(* Logix 5000 project; controller Test vendor 1 type 14 code 167 rev 35.11; software revision 35.00 *)

TASK MainTask (continuous, watchdog 500 ms) : MainProgram

MODULES
   Local : vendor 1 type 14 code 167 (ICP 0, rev 35.11)
END_MODULES

TYPE CMoDateTime :   // Date and Time Structure
STRUCT
   RawDateTime : DINT[7];   // Platform-native wall clock data
   Year : DINT;
   Month : DINT;   // 1-12
   Day : DINT;   // 1-31
   Hour : DINT;   // 0-23
   Minute : DINT;   // 0-59
   Second : DINT;   // 0-59
   MicroSecond : DINT;   // 0-999999
   IsLocal : BOOL;   // TRUE = local time, FALSE = UTC
END_STRUCT
END_TYPE

TYPE CMoDateTimeString :   // HMI-Readable Date/Time Strings
STRUCT
   TimeString : CMoString28;   // HH:MM:SS
   DateString : CMoString28;   // YYYY-MM-DD
   HMIString : CMoString28;   // YYYY-MM-DD HH:MM:SS
END_STRUCT
END_TYPE

TYPE CMoFramework :   // Shared System Context - one per PLC
STRUCT
   AnyAudibleOn : BOOL;   // Audible alarm active
   AnyAudibleOnLastScan : BOOL;   // Scratch
   AnyAlarmActive : BOOL;   // Alarm active
   AnyAlarmActiveLastScan : BOOL;   // Scratch
   AnyWarningActive : BOOL;   // Warning active
   AnyWarningActiveLastScan : BOOL;   // Scratch
   AnyFaultActive : BOOL;   // Fault active
   AnyFaultActiveLastScan : BOOL;   // Scratch
   AnyCriticalActive : BOOL;   // Critical active
   AnyCriticalActiveLastScan : BOOL;   // Scratch
   AnySimulationOn : BOOL;   // Sim active
   AnySimulationOnLastScan : BOOL;   // Scratch
   AnyHandOn : BOOL;   // Hand active
   AnyHandOnLastScan : BOOL;   // Scratch
   SilenceCmd : BOOL;   // HMI silence (momentary)
   GlobalAlmRstCmd : BOOL;   // HMI global reset (momentary)
   GlobalAlmRstEn : BOOL;   // Enable global reset
   SimulationEnabled : BOOL;   // Master sim enable
   EmulationEnabled : BOOL;   // Emulated controller
   MaintenanceEnabled : BOOL;   // Enables Hand mode
   Tick100ms : BOOL;   // 100ms tick
   Tick1s : BOOL;   // 1s tick
   Tick10s : BOOL;   // 10s tick
   Blink100ms : BOOL;   // 100ms blinker
   Blink250ms : BOOL;   // 250ms blinker
   Blink500ms : BOOL;   // 500ms blinker
   Blink1s : BOOL;   // 1s blinker
   Blink2s : BOOL;   // 2s blinker
   InhibitAlarms : BOOL;   // Corporate alarm inhibit
   AlwaysTrue : BOOL;   // Constant TRUE
   AlwaysFalse : BOOL;   // Constant FALSE
   ApplicationCount : DINT;   // AOI instance count
   AlarmCount : INT;   // Active alarm count
   TempAlarmCount : INT;   // Scratch
   FreeRunningTimer : DINT;   // Free-running ms counter
   LastRandomSeed : DINT;   // Random seed
   Random : REAL;   // Random 0.0-1.0
   CycleTime : REAL;   // Scan time (ms)
   InhibitAlarmGroups : DINT[16];   // Per-group inhibit (512 groups)
   CurrentUTCDateTime : CMoDateTime;   // UTC time
   CurrentLocalDateTime : CMoDateTime;   // Local time
   CurrentUTCString : CMoDateTimeString;   // UTC strings
   CurrentLocalString : CMoDateTimeString;   // Local strings
   NotUsedDI : CMoHALDigitalInput;   // Spare DI
   NotUsedDO : CMoHALDigitalOutput;   // Spare DO
   ModuleStatusMinInterval : DINT;   // ms between module checks
   ModuleStatusRandomDistribution : DINT;   // ms random spread
   ModuleStatusGraceTime : DINT;   // ms before module lost
END_STRUCT
END_TYPE

TYPE CMoHALDigitalInput :   // Digital Input HAL - Business logic reads .Value only
STRUCT
   Input : BOOL;   // Raw hardware input
   QualityInput : BOOL;   // Hardware health (TRUE = good)
   SimInput : BOOL;   // Simulation input (twin/test)
   EnableSimulation : BOOL;   // Enable simulation for this point
   SimulationIsActive : BOOL;   // Computed: EnableSimulation AND Framework.SimulationEnabled
   HandValue : BOOL;   // Manual override value (HMI)
   EnableHand : BOOL;   // Enable hand mode
   HandIsActive : BOOL;   // Computed: EnableHand AND Framework.MaintenanceEnabled
   Value : BOOL;   // THE OUTPUT: conditioned, filtered, mode-selected
   Inverted : BOOL;   // Invert input polarity
   BadQualityValue : BOOL;   // Value when quality is bad
   EnableDelay : BOOL;   // Enable debounce filtering
   IsSpare : BOOL;   // Mark as spare
   InFilterOnTimeMsec : DINT;   // On-delay debounce (ms)
   InFilterOffTimeMsec : DINT;   // Off-delay debounce (ms)
   PointQuality : BOOL;   // Computed quality
   RisingEdge : BOOL;   // One-shot on Value 0->1
   FallingEdge : BOOL;   // One-shot on Value 1->0
   Name : CMoString28;   // Human-readable tag name
END_STRUCT
END_TYPE

TYPE CMoHALDigitalOutput :   // Digital Output HAL - Business logic writes .Value
STRUCT
   Output : BOOL;   // Physical output
   QualityInput : BOOL;   // Hardware health (TRUE = good)
   SimOutput : BOOL;   // Shadow output for twin
   EnableSimulation : BOOL;   // Enable simulation
   SimulationIsActive : BOOL;   // Computed
   HandValue : BOOL;   // Manual override value
   EnableHand : BOOL;   // Enable hand mode
   HandIsActive : BOOL;   // Computed
   Value : BOOL;   // Business logic command
   Inverted : BOOL;   // Invert output polarity
   BadQualityValue : BOOL;   // Value when quality is bad
   IsSpare : BOOL;   // Mark as spare
   PointQuality : BOOL;   // Computed quality
   Name : CMoString28;   // Human-readable tag name
END_STRUCT
END_TYPE

TYPE CMoInterlock :   // Interlock: 16 AND conditions, first-out, per-condition bypass
STRUCT
   PointCount : INT;   // Number of active conditions (1-16)
   Condition : BOOL[32];   // Condition inputs
   Bypass : BOOL[32];   // Per-condition bypass (HMI)
   OK : BOOL;   // All conditions met or bypassed
   InBypass : BOOL;   // At least one bypassed
   BypassAlarm : BOOL;   // Operating with bypass
   FirstOut : INT;   // First faulted condition index (-1=none)
   ConditionMet : BOOL[32];   // Condition OR bypass
   ConditionFaulted : BOOL[32];   // Failed AND not bypassed
   Name : CMoString28;   // Interlock name
   ConditionName : CMoString28[16];   // Per-condition labels
END_STRUCT
END_TYPE

TYPE CMoString28 :
STRUCT
   LEN : DINT;
   DATA : SINT[28];
END_STRUCT
END_TYPE

ADD_ON_INSTRUCTION CMoAlarm   (* revision 1.0 *)
// Alarm Monitor
// Help:
// Trigger, delay, reset, severity, group inhibit, silencing, occurrence counting.
VAR_IN_OUT
   Framework : CMoFramework; {required}   // System context
END_VAR
VAR_INPUT
   Trigger : BOOL;   // Condition to monitor
   EnableAlarm : BOOL := 1;   // Enable this alarm
   AlarmOnTrue : BOOL := 1;   // Trigger=1 alarms
   AutoReset : BOOL;   // Auto-clear
   Delay : DINT;   // ms before activating
   GroupNo : DINT;   // Alarm group 0-511
   ID : INT;   // Alarm ID 1-9023
   IsWarning : BOOL;   // Warning severity
   IsFault : BOOL;   // Fault severity
   IsCritical : BOOL;   // Critical severity
   EnableAudio : BOOL;   // Enable audible
   SystemResetEnable : BOOL := 1;   // Allow global reset
   Reset : BOOL;   // Manual reset
   Inhibit : BOOL;   // Per-alarm inhibit
   CountPreset : DINT;   // Count threshold
   CountReset : BOOL;   // Reset counter
END_VAR
VAR_OUTPUT
   AlarmActive : BOOL; {access Read Only}   // Alarm is active
   InhibitActive : BOOL; {access Read Only}   // Currently inhibited
   AlarmCount : DINT; {access Read Only}   // Activation count
   CountExceeded : BOOL; {access Read Only}   // Count >= preset
   AlarmSilenced : BOOL; {access Read Only}   // Active but silenced
END_VAR
VAR
   AlarmTimer : FBD_TIMER; {access None}
   IntGroupNo : DINT; {access None}
   IntID : DINT; {access None}
   IntReset : BOOL; {access None}
   TriggerCondition : BOOL; {access None}
   PrevAlarmActive : BOOL; {access None}
END_VAR

ROUTINE Logic   (* structured text *)
   // =============================================================================
   // CMoAlarm — Alarm Monitor
   // CMo Library v1.0
   // =============================================================================
   // Monitors a trigger condition and manages alarm lifecycle.
   // Supports configurable trigger polarity, delay before activation,
   // auto/manual reset, occurrence counting with threshold,
   // severity classification (Warning/Fault/Critical), group-based
   // inhibit, and HMI silencing.
   // =============================================================================
   
   IF GroupNo >= 0 AND GroupNo <= 511 THEN IntGroupNo := GroupNo; ELSE IntGroupNo := 0; END_IF;
   IF ID >= 1 AND ID <= 9023 THEN IntID := ID; ELSE IntID := 0; END_IF;
   IF CountReset THEN AlarmCount := 0; CountReset := 0; END_IF;
   InhibitActive := NOT EnableAlarm OR Inhibit OR Framework.InhibitAlarms;
   IntReset := AutoReset OR Reset OR (SystemResetEnable AND Framework.GlobalAlmRstEn AND Framework.GlobalAlmRstCmd);
   IF AlarmOnTrue THEN TriggerCondition := Trigger; ELSE TriggerCondition := NOT Trigger; END_IF;
   
   IF IntID <> 0 THEN
       AlarmTimer.PRE := Delay;
       AlarmTimer.TimerEnable := (NOT InhibitActive AND TriggerCondition) OR (AlarmActive AND NOT IntReset);
       TONR(AlarmTimer);
       AlarmActive := AlarmTimer.DN;
       IF NOT AlarmTimer.TimerEnable THEN
           AlarmTimer.Reset := 1; TONR(AlarmTimer); AlarmTimer.Reset := 0;
       END_IF;
   ELSE
       AlarmActive := 0;
   END_IF;
   
   IF AlarmActive AND NOT PrevAlarmActive THEN AlarmCount := AlarmCount + 1; END_IF;
   IF AlarmActive THEN
       IF Framework.SilenceCmd OR AlarmSilenced THEN AlarmSilenced := 1; END_IF;
   ELSE AlarmSilenced := 0;
   END_IF;
   
   IF AlarmActive THEN
       Framework.TempAlarmCount := Framework.TempAlarmCount + 1;
       Framework.AnyAlarmActiveLastScan := 1;
       IF NOT AlarmSilenced THEN
           IF EnableAudio THEN Framework.AnyAudibleOnLastScan := 1; END_IF;
           IF IsWarning THEN Framework.AnyWarningActiveLastScan := 1; END_IF;
           IF IsFault THEN Framework.AnyFaultActiveLastScan := 1; END_IF;
           IF IsCritical THEN Framework.AnyCriticalActiveLastScan := 1; END_IF;
       END_IF;
   END_IF;
   
   IF CountPreset > 0 AND AlarmCount >= CountPreset THEN CountExceeded := 1; ELSE CountExceeded := 0; END_IF;
   Reset := 0;
   PrevAlarmActive := AlarmActive;
END_ROUTINE
END_ADD_ON_INSTRUCTION

ADD_ON_INSTRUCTION CMoDateTimeToString   (* revision 1.0 *)
// Format DateTime for HMI Display
// Help:
// Converts CMoDateTime into zero-padded strings.
VAR_IN_OUT
   DateTime : CMoDateTime; {required}   // Input DateTime
   DateTimeString : CMoDateTimeString; {required}   // Output formatted strings
END_VAR
VAR
   sYear : CMoString28; {access None}
   sMonth : CMoString28; {access None}
   sDay : CMoString28; {access None}
   sHour : CMoString28; {access None}
   sMinute : CMoString28; {access None}
   sSecond : CMoString28; {access None}
   sTemp : CMoString28; {access None}
   sZero : CMoString28; {access None}
   sColon : CMoString28; {access None}
   sDash : CMoString28; {access None}
   sBlank : CMoString28; {access None}
END_VAR

ROUTINE Logic   (* structured text *)
   // =============================================================================
   // CMoDateTimeToString — Format DateTime for HMI Display
   // CMo Library v1.0
   // =============================================================================
   // Converts CMoDateTime fields into zero-padded human-readable strings:
   //   TimeString: "HH:MM:SS"
   //   DateString: "YYYY-MM-DD"
   //   HMIString:  "YYYY-MM-DD HH:MM:SS"
   //
   // Uses DTOS for DINT-to-string conversion.
   // =============================================================================
   
   DTOS(DateTime.Year, sYear);
   sZero := '0';
   sColon := ':';
   sDash := '-';
   sBlank := ' ';
   IF DateTime.Month < 10 THEN
       DTOS(DateTime.Month, sTemp);
       CONCAT(sZero, sTemp, sMonth);
   ELSE
       DTOS(DateTime.Month, sMonth);
   END_IF;
   
   IF DateTime.Day < 10 THEN
       DTOS(DateTime.Day, sTemp);
       CONCAT(sZero, sTemp, sDay);
   ELSE
       DTOS(DateTime.Day, sDay);
   END_IF;
   
   IF DateTime.Hour < 10 THEN
       DTOS(DateTime.Hour, sTemp);
       CONCAT(sZero, sTemp, sHour);
   ELSE
       DTOS(DateTime.Hour, sHour);
   END_IF;
   
   IF DateTime.Minute < 10 THEN
       DTOS(DateTime.Minute, sTemp);
       CONCAT(sZero, sTemp, sMinute);
   ELSE
       DTOS(DateTime.Minute, sMinute);
   END_IF;
   
   IF DateTime.Second < 10 THEN
       DTOS(DateTime.Second, sTemp);
       CONCAT(sZero, sTemp, sSecond);
   ELSE
       DTOS(DateTime.Second, sSecond);
   END_IF;
   
   // Build TimeString: "HH:MM:SS"
   
   CONCAT(sHour, sColon, sTemp);
   CONCAT(sTemp, sMinute, sTemp);
   CONCAT(sTemp, sColon, sTemp);
   CONCAT(sTemp, sSecond, DateTimeString.TimeString);
   
   // Build DateString: "YYYY-MM-DD"
   CONCAT(sYear, sDash, sTemp);
   CONCAT(sTemp, sMonth, sTemp);
   CONCAT(sTemp, sDash, sTemp);
   CONCAT(sTemp, sDay, DateTimeString.DateString);
   
   // Build HMIString: "YYYY-MM-DD HH:MM:SS"
   CONCAT(DateTimeString.DateString, sBlank, sTemp);
   CONCAT(sTemp, DateTimeString.TimeString, DateTimeString.HMIString);
END_ROUTINE
END_ADD_ON_INSTRUCTION

ADD_ON_INSTRUCTION CMoDiffTime   (* revision 1.0 *)
// DateTime Subtraction with Carry Propagation
// Help:
// Computes EndTime - StartTime with carry propagation.
VAR_IN_OUT
   StartTime : CMoDateTime; {required}   // Start time
   EndTime : CMoDateTime; {required}   // End time
   Result : CMoDateTime; {required}   // Difference result
END_VAR
VAR_OUTPUT
   TotalSeconds : DINT; {access Read Only}   // Approximate total seconds
   TotalMicroseconds : DINT; {access Read Only}   // Remainder microseconds
END_VAR
VAR
   a : DINT; {access None}
   y : DINT; {access None}
   m : DINT; {access None}
   jdnStart : DINT; {access None}
   jdnEnd : DINT; {access None}
   diffDays : DINT; {access None}
   diffUs : DINT; {access None}
   diffSec : DINT; {access None}
   diffMin : DINT; {access None}
   diffHr : DINT; {access None}
END_VAR

ROUTINE Logic   (* structured text *)
   // =============================================================================
   // CMoDiffTime — DateTime Subtraction via Julian Day Number
   // CMo Library v1.0 — Rockwell
   // =============================================================================
   // Computes (EndTime - StartTime) using Julian Day Number conversion.
   // Converts both dates to JDN (integer day count), subtracts, then
   // handles sub-day time remainder with borrow propagation.
   //
   // This is mathematically correct for all valid dates regardless of
   // month lengths, leap years, or century boundaries.
   //
   // Usage:
   //   CMoDiffTime(fbDiff, tStart, tEnd, tResult);
   //   elapsed := fbDiff.TotalSeconds;
   // =============================================================================
   
   // JDN for StartTime
   a := (14 - StartTime.Month) / 12;
   y := StartTime.Year + 4800 - a;
   m := StartTime.Month + 12 * a - 3;
   jdnStart := StartTime.Day + (153 * m + 2) / 5 + 365 * y + y / 4 - y / 100 + y / 400 - 32045;
   
   // JDN for EndTime
   a := (14 - EndTime.Month) / 12;
   y := EndTime.Year + 4800 - a;
   m := EndTime.Month + 12 * a - 3;
   jdnEnd := EndTime.Day + (153 * m + 2) / 5 + 365 * y + y / 4 - y / 100 + y / 400 - 32045;
   
   // Day difference
   diffDays := jdnEnd - jdnStart;
   
   // Sub-day difference with borrow propagation
   diffUs := EndTime.MicroSecond - StartTime.MicroSecond;
   IF diffUs < 0 THEN
       diffUs := diffUs + 1000000;
       diffSec := -1;
   ELSE
       diffSec := 0;
   END_IF;
   
   diffSec := diffSec + EndTime.Second - StartTime.Second;
   IF diffSec < 0 THEN
       diffSec := diffSec + 60;
       diffMin := -1;
   ELSE
       diffMin := 0;
   END_IF;
   
   diffMin := diffMin + EndTime.Minute - StartTime.Minute;
   IF diffMin < 0 THEN
       diffMin := diffMin + 60;
       diffHr := -1;
   ELSE
       diffHr := 0;
   END_IF;
   
   diffHr := diffHr + EndTime.Hour - StartTime.Hour;
   IF diffHr < 0 THEN
       diffHr := diffHr + 24;
       diffDays := diffDays - 1;
   END_IF;
   
   // Populate result
   Result.Year := 0;
   Result.Month := 0;
   Result.Day := diffDays;
   Result.Hour := diffHr;
   Result.Minute := diffMin;
   Result.Second := diffSec;
   Result.MicroSecond := diffUs;
   Result.IsLocal := 0;
   
   // Convenience totals
   TotalSeconds := diffSec + (diffMin * 60) + (diffHr * 3600) + (diffDays * 86400);
   TotalMicroseconds := diffUs;
END_ROUTINE
END_ADD_ON_INSTRUCTION

ADD_ON_INSTRUCTION CMoDigitalInput   (* revision 1.0 *)
// Digital Input Signal Conditioning
// Help:
// Mode select, inversion, debounce, quality gating, edge detection. Reads .Value only.
VAR_IN_OUT
   HAL : CMoHALDigitalInput; {required}   // HAL Interface
END_VAR
VAR_INPUT
   DeviceInput : BOOL; {required}   // Raw hardware input
   QualityInput : BOOL; {required}   // Module health
END_VAR
VAR_IN_OUT
   Framework : CMoFramework; {required}   // System context
END_VAR
VAR
   ConditionedInput : BOOL; {access None}
   DebouncedValue : BOOL; {access None}
   OnDelayTimer : FBD_TIMER; {access None}
   OffDelayTimer : FBD_TIMER; {access None}
   PrevValue : BOOL; {access None}
   FirstScan : BOOL := 1; {access None}
   ReSync : BOOL; {access None}
   NoFilterNeeded : BOOL; {access None}
END_VAR

ROUTINE Logic   (* structured text *)
   // =============================================================================
   // CMoDigitalInput — Digital Input Signal Conditioning
   // CMo Library v1.0
   // =============================================================================
   // Takes a raw hardware input and produces a conditioned .Value through:
   //   1. Mode determination (Normal / Simulation / Hand)
   //   2. Quality evaluation (hardware health, sim, spare)
   //   3. Mode selection + polarity inversion
   //   4. Debounce filtering (configurable on/off delay with resync)
   //   5. Hand value bumpless transfer
   //   6. Quality gating (bad quality -> configurable fallback)
   //   7. Edge detection (RisingEdge / FallingEdge one-shot pulses)
   //
   // Business logic reads .Value only.
   // =============================================================================
   
   // Mode determination
   HAL.HandIsActive := HAL.EnableHand AND Framework.MaintenanceEnabled;
   IF HAL.HandIsActive THEN Framework.AnyHandOnLastScan := 1; END_IF;
   HAL.SimulationIsActive := HAL.EnableSimulation AND Framework.SimulationEnabled;
   IF HAL.SimulationIsActive THEN Framework.AnySimulationOnLastScan := 1; END_IF;
   
   // Point quality
   IF HAL.IsSpare THEN HAL.PointQuality := 1;
   ELSIF HAL.SimulationIsActive THEN HAL.PointQuality := 1;
   ELSE HAL.QualityInput := QualityInput; HAL.PointQuality := QualityInput;
   END_IF;
   
   // Latch raw input
   HAL.Input := DeviceInput;
   
   // Mode selection + inversion
   IF HAL.SimulationIsActive THEN
       IF HAL.Inverted THEN ConditionedInput := NOT HAL.SimInput;
       ELSE ConditionedInput := HAL.SimInput; END_IF;
   ELSE
       IF HAL.Inverted THEN ConditionedInput := NOT HAL.Input;
       ELSE ConditionedInput := HAL.Input; END_IF;
   END_IF;
   
   // Debounce filter
   IF NOT HAL.EnableDelay THEN
       DebouncedValue := ConditionedInput; ReSync := 1;
   ELSE
       IF HAL.InFilterOnTimeMsec < 0 THEN HAL.InFilterOnTimeMsec := 0; END_IF;
       IF HAL.InFilterOffTimeMsec < 0 THEN HAL.InFilterOffTimeMsec := 0; END_IF;
       OnDelayTimer.PRE := HAL.InFilterOnTimeMsec;
       OnDelayTimer.TimerEnable := ConditionedInput;
       TONR(OnDelayTimer);
       OffDelayTimer.PRE := HAL.InFilterOffTimeMsec;
       OffDelayTimer.TimerEnable := NOT ConditionedInput;
       TONR(OffDelayTimer);
       IF ReSync THEN
           IF (DebouncedValue AND OnDelayTimer.DN) OR (NOT DebouncedValue AND NOT OnDelayTimer.DN) THEN ReSync := 0; END_IF;
       END_IF;
       IF ReSync OR HAL.IsSpare THEN DebouncedValue := ConditionedInput;
       ELSIF OnDelayTimer.DN THEN DebouncedValue := 1;
           OffDelayTimer.Reset := 1; TONR(OffDelayTimer); OffDelayTimer.Reset := 0;
       END_IF;
       IF NOT ConditionedInput AND OffDelayTimer.DN THEN DebouncedValue := 0;
           OnDelayTimer.Reset := 1; TONR(OnDelayTimer); OnDelayTimer.Reset := 0;
       END_IF;
   END_IF;
   
   // Hand value tracking (bumpless transfer)
   IF NOT HAL.HandIsActive THEN HAL.HandValue := HAL.Value; END_IF;
   
   // Final value with quality gating
   IF HAL.PointQuality THEN
       IF HAL.HandIsActive THEN HAL.Value := HAL.HandValue;
       ELSE HAL.Value := DebouncedValue; END_IF;
   ELSE HAL.Value := HAL.BadQualityValue;
   END_IF;
   
   // Edge detection
   IF FirstScan THEN
       PrevValue := HAL.Value; HAL.RisingEdge := 0; HAL.FallingEdge := 0; FirstScan := 0;
   ELSE
       HAL.RisingEdge := HAL.Value AND NOT PrevValue;
       HAL.FallingEdge := NOT HAL.Value AND PrevValue;
       PrevValue := HAL.Value;
   END_IF;
END_ROUTINE
END_ADD_ON_INSTRUCTION

ADD_ON_INSTRUCTION CMoDigitalOutput   (* revision 1.0 *)
// Digital Output Signal Conditioning
// Help:
// Mode select, inversion, hand, sim gating. Writes .Value, twin reads .SimOutput.
VAR_IN_OUT
   HAL : CMoHALDigitalOutput; {required}   // HAL Interface
END_VAR
VAR_INPUT
   QualityInput : BOOL; {required}   // Module health
END_VAR
VAR_OUTPUT
   DeviceOutput : BOOL; {access Read Only, visible}   // Physical output
END_VAR
VAR_IN_OUT
   Framework : CMoFramework; {required}   // System context
END_VAR
VAR
   ConditionedOutput : BOOL; {access None}
   OutputWithHand : BOOL; {access None}
END_VAR

ROUTINE Logic   (* structured text *)
   // =============================================================================
   // CMoDigitalOutput — Digital Output Signal Conditioning
   // CMo Library v1.0
   // =============================================================================
   // Takes .Value written by business logic and produces a conditioned
   // physical output through:
   //   1. Mode determination (Normal / Simulation / Hand)
   //   2. Quality evaluation (hardware health, sim, spare)
   //   3. Polarity inversion
   //   4. Hand value bumpless transfer
   //   5. Hand mode selection
   //   6. Simulation gating (suppress physical output, capture to .SimOutput)
   //
   // In simulation mode: DeviceOutput is suppressed. The digital twin
   // reads .SimOutput to see what business logic commanded.
   //
   // Usage:
   //   CMoDigitalOutput(fbOutput, HAL, Module2_Status.Running, Framework);
   //   Module2:O.Data[0] := fbOutput.DeviceOutput;
   // =============================================================================
   
   HAL.HandIsActive := HAL.EnableHand AND Framework.MaintenanceEnabled AND NOT HAL.IsSpare;
   IF HAL.HandIsActive THEN Framework.AnyHandOnLastScan := 1; END_IF;
   HAL.SimulationIsActive := HAL.EnableSimulation AND Framework.SimulationEnabled;
   IF HAL.SimulationIsActive THEN Framework.AnySimulationOnLastScan := 1; END_IF;
   IF HAL.IsSpare THEN HAL.PointQuality := 1;
   ELSIF HAL.SimulationIsActive THEN HAL.PointQuality := 1;
   ELSE HAL.QualityInput := QualityInput; HAL.PointQuality := QualityInput;
   END_IF;
   IF NOT HAL.IsSpare THEN
       IF HAL.Inverted THEN ConditionedOutput := NOT HAL.Value;
       ELSE ConditionedOutput := HAL.Value; END_IF;
   ELSE ConditionedOutput := 0;
   END_IF;
   IF NOT HAL.HandIsActive THEN HAL.HandValue := HAL.Value; END_IF;
   IF HAL.HandIsActive THEN OutputWithHand := HAL.HandValue;
   ELSE OutputWithHand := ConditionedOutput; END_IF;
   IF HAL.SimulationIsActive THEN DeviceOutput := 0;
   ELSE DeviceOutput := OutputWithHand; END_IF;
   HAL.SimOutput := OutputWithHand;
   HAL.Output := DeviceOutput;
END_ROUTINE
END_ADD_ON_INSTRUCTION

ADD_ON_INSTRUCTION CMoElapsedTime   (* revision 1.0 *)
// Elapsed Time Measurement
// Help:
// Measures elapsed time between Start and Stop rising edges.
VAR_INPUT
   Start : BOOL; {required}   // Begin measurement
   Stop : BOOL; {required}   // End measurement
   Reset : BOOL; {required}   // Clear measurement
END_VAR
VAR_OUTPUT
   ElapsedMs : REAL; {access Read Only}   // Result in ms
   Running : BOOL; {access Read Only}   // TRUE while measuring
END_VAR
VAR
   PrevStart : BOOL; {access None}
   PrevStop : BOOL; {access None}
   tmRun : FBD_TIMER; {access None}
   Capturing : BOOL; {access None}
END_VAR

ROUTINE Logic   (* structured text *)
   // =============================================================================
   // CMoElapsedTime — Elapsed Time Measurement
   // CMo Library v1.0
   // =============================================================================
   // Measures elapsed time between Start and Stop rising edges.
   // Uses TONR timer internally for millisecond-resolution measurement.
   // Live readout available via ElapsedMs while Running is TRUE.
   //
   // Usage:
   //   CMoElapsedTime(myTimer, TRUE, FALSE, FALSE);  // Start
   //   CMoElapsedTime(myTimer, FALSE, TRUE, FALSE);  // Stop
   //   result := myTimer.ElapsedMs;
   //   CMoElapsedTime(myTimer, FALSE, FALSE, TRUE);  // Reset
   // =============================================================================
   
   IF Reset THEN
       ElapsedMs := 0.0;
       Running := 0;
       Capturing := 0;
       tmRun.Reset := 1;
       TONR(tmRun);
       tmRun.Reset := 0;
       TND();
   END_IF;
   
   IF Start AND NOT PrevStart THEN
       Capturing := 1;
       Running := 1;
       tmRun.Reset := 1;
       TONR(tmRun);
       tmRun.Reset := 0;
       tmRun.PRE := 2147483647;
   END_IF;
   PrevStart := Start;
   
   IF Capturing THEN
       tmRun.TimerEnable := 1;
       TONR(tmRun);
       ElapsedMs := tmRun.ACC;
   END_IF;
   
   IF Stop AND NOT PrevStop AND Capturing THEN
       ElapsedMs := tmRun.ACC;
       tmRun.TimerEnable := 0;
       Capturing := 0;
       Running := 0;
   END_IF;
   PrevStop := Stop;
END_ROUTINE
END_ADD_ON_INSTRUCTION

ADD_ON_INSTRUCTION CMoEvalInterlock   (* revision 1.0 *)
// Interlock Evaluation
// Help:
// Up to 16 AND conditions, first-out tracking, per-condition bypass.
VAR_IN_OUT
   Ilk : CMoInterlock; {required}   // Interlock structure
END_VAR
VAR
   i : DINT; {access None}
   AllMet : BOOL; {access None}
   AnyBypassed : BOOL; {access None}
   FirstDropped : INT; {access None}
   PrevOK : BOOL; {access None}
END_VAR

ROUTINE Logic   (* structured text *)
   // =============================================================================
   // CMoEvalInterlock — Interlock Evaluation
   // CMo Library v1.0
   // =============================================================================
   // Evaluates up to 16 AND conditions with first-out tracking
   // and per-condition bypass. All active conditions must be TRUE
   // (or bypassed) for .OK to be TRUE.
   //
   // FirstOut latches the index of the first faulted condition on
   // the OK->NOT OK transition (root cause analysis from HMI).
   //
   // Usage:
   //   Ilk.Condition[0] := EStop.Value;
   //   Ilk.Condition[1] := GuardDoor.Value;
   //   CMoEvalInterlock(fbInterlock, MyInterlock);
   //   IF MyInterlock.OK THEN ... END_IF;
   // =============================================================================
   
   IF Ilk.PointCount < 1 THEN Ilk.PointCount := 1; ELSIF Ilk.PointCount > 16 THEN Ilk.PointCount := 16; END_IF;
   AllMet := 1; AnyBypassed := 0; FirstDropped := -1;
   FOR i := 0 TO Ilk.PointCount - 1 DO
       Ilk.ConditionMet[i] := Ilk.Condition[i] OR Ilk.Bypass[i];
       Ilk.ConditionFaulted[i] := NOT Ilk.Condition[i] AND NOT Ilk.Bypass[i];
       IF Ilk.Bypass[i] THEN AnyBypassed := 1; END_IF;
       IF Ilk.ConditionFaulted[i] AND FirstDropped = -1 THEN FirstDropped := i; END_IF;
       IF NOT Ilk.ConditionMet[i] THEN AllMet := 0; END_IF;
   END_FOR;
   FOR i := Ilk.PointCount TO 15 DO
       Ilk.ConditionMet[i] := 1; Ilk.ConditionFaulted[i] := 0;
   END_FOR;
   PrevOK := Ilk.OK;
   Ilk.OK := AllMet; Ilk.InBypass := AnyBypassed; Ilk.BypassAlarm := AnyBypassed;
   IF NOT Ilk.OK AND PrevOK THEN Ilk.FirstOut := FirstDropped;
   ELSIF Ilk.OK THEN Ilk.FirstOut := -1; END_IF;
END_ROUTINE
END_ADD_ON_INSTRUCTION

ADD_ON_INSTRUCTION CMoGetLocalDateTime   (* revision 1.0 *)
// Read Local System Time (Rockwell)
// Help:
// Reads PLC wall clock via GSV WallClockTime into CMoDateTime.
VAR_IN_OUT
   DateTime : CMoDateTime; {required}   // Output DateTime structure
END_VAR

ROUTINE Logic   (* structured text *)
   // =============================================================================
   // CMoGetLocalDateTime — Read Local System Time (Rockwell)
   // CMo Library v1.0
   // =============================================================================
   // Reads PLC wall clock via GSV WallClockTime into CMoDateTime.
   // GSV WallClockTime returns local time as DINT[7]:
   //   [Year, Month, Day, Hour, Minute, Second, MicroSecond]
   //
   // Must be called cyclically. Called internally by CMoMainRuntime.
   //
   // Usage:
   //   CMoGetLocalDateTime(fbLocal, Framework.CurrentLocalDateTime);
   // =============================================================================
   
   GSV(WallClockTime,,LocalDateTime,DateTime.RawDateTime[0]);
   DateTime.Year := DateTime.RawDateTime[0];
   DateTime.Month := DateTime.RawDateTime[1];
   DateTime.Day := DateTime.RawDateTime[2];
   DateTime.Hour := DateTime.RawDateTime[3];
   DateTime.Minute := DateTime.RawDateTime[4];
   DateTime.Second := DateTime.RawDateTime[5];
   DateTime.MicroSecond := DateTime.RawDateTime[6];
   DateTime.IsLocal := 1;
END_ROUTINE
END_ADD_ON_INSTRUCTION

ADD_ON_INSTRUCTION CMoGetUTCDateTime   (* revision 1.0 *)
// Read UTC System Time (Rockwell)
// Help:
// Reads PLC wall clock via GSV WallClockTime. Set controller clock to UTC for true UTC.
VAR_IN_OUT
   DateTime : CMoDateTime; {required}   // Output DateTime structure
END_VAR

ROUTINE Logic   (* structured text *)
   // =============================================================================
   // CMoGetUTCDateTime — Read UTC System Time (Rockwell)
   // CMo Library v1.0
   // =============================================================================
   // Reads PLC wall clock via GSV WallClockTime.
   // Note: Rockwell GSV returns local time. For true UTC,
   // configure controller clock to UTC or apply offset.
   //
   // Called internally by CMoMainRuntime.
   //
   // Usage:
   //   CMoGetUTCDateTime(fbUTC, Framework.CurrentUTCDateTime);
   // =============================================================================
   
   GSV(WallClockTime,,DateTime,DateTime.RawDateTime[0]);
   DateTime.Year := DateTime.RawDateTime[0];
   DateTime.Month := DateTime.RawDateTime[1];
   DateTime.Day := DateTime.RawDateTime[2];
   DateTime.Hour := DateTime.RawDateTime[3];
   DateTime.Minute := DateTime.RawDateTime[4];
   DateTime.Second := DateTime.RawDateTime[5];
   DateTime.MicroSecond := DateTime.RawDateTime[6];
   DateTime.IsLocal := 0;
END_ROUTINE
END_ADD_ON_INSTRUCTION

ADD_ON_INSTRUCTION CMoMainRuntime   (* revision 1.0 *)
// System Heartbeat - call ONCE per scan, FIRST in the task
// Help:
// Scan time, ticks, blinkers, alarm rollups, random, date/time. Calls CMoElapsedTime, CMoRandom, CMoGetLocalDateTime, CMoGetUTCDateTime, CMoDateTimeToString.
VAR_IN_OUT
   Framework : CMoFramework; {required}   // Shared system context
END_VAR
VAR
   tmTick100ms : FBD_TIMER; {access None}
   tmTick1s : FBD_TIMER; {access None}
   tmTick10s : FBD_TIMER; {access None}
   tmBlink100ms : FBD_TIMER; {access None}
   tmBlink250ms : FBD_TIMER; {access None}
   tmBlink500ms : FBD_TIMER; {access None}
   tmBlink1s : FBD_TIMER; {access None}
   tmBlink2s : FBD_TIMER; {access None}
   bState100ms : BOOL; {access None}
   bState250ms : BOOL; {access None}
   bState500ms : BOOL; {access None}
   bState1s : BOOL; {access None}
   bState2s : BOOL; {access None}
   bScanRunning : BOOL; {access None}
   fbScanTime : CMoElapsedTime; {access None}
   fbRandom : CMoRandom := (Seed := 48271); {access None}
   fbGetLocal : CMoGetLocalDateTime; {access None}
   fbGetUTC : CMoGetUTCDateTime; {access None}
   fbLocalToStr : CMoDateTimeToString; {access None}
   fbUTCToStr : CMoDateTimeToString; {access None}
END_VAR

ROUTINE Logic   (* structured text *)
   // =============================================================================
   // CMoMainRuntime — System Heartbeat
   // CMo Library v1.0
   // =============================================================================
   // Call ONCE per scan, FIRST in the task. Responsible for:
   //   - Measuring scan cycle time (via CMoElapsedTime)
   //   - Generating tick timers (100ms, 1s, 10s)
   //   - Generating blinker signals (100ms, 250ms, 500ms, 1s, 2s)
   //   - Latching LastScan accumulators into final alarm/sim/hand rollups
   //   - Resetting LastScan accumulators for the new scan
   //   - Generating random number (via CMoRandom)
   //   - Updating local and UTC date/time with formatted strings
   //   - Setting constants (AlwaysTrue, AlwaysFalse)
   //   - Incrementing free-running timer
   //
   // The LastScan pattern:
   //   MainRuntime resets all *LastScan fields at start of scan.
   //   Individual CMoAlarm/CMoDigitalInput AOIs SET them during the scan.
   //   MainRuntime copies LastScan -> final at the NEXT call.
   //   This eliminates execution order dependencies.
   //
   // Usage:
   //   CMoMainRuntime(fbRuntime, Framework);  // first line of MainRoutine
   // =============================================================================
   
   // Scan time measurement
   IF bScanRunning THEN
       CMoElapsedTime(fbScanTime,0,1,0);
       Framework.CycleTime := fbScanTime.ElapsedMs;
       CMoElapsedTime(fbScanTime,0,0,1);
       CMoElapsedTime(fbScanTime,1,0,0);
   ELSE
       CMoElapsedTime(fbScanTime,1,0,0);
       bScanRunning := 1;
   END_IF;
   
   // Latch previous scan accumulators
   Framework.AnyAudibleOn := Framework.AnyAudibleOnLastScan;
   Framework.AnyAlarmActive := Framework.AnyAlarmActiveLastScan;
   Framework.AnyWarningActive := Framework.AnyWarningActiveLastScan;
   Framework.AnyFaultActive := Framework.AnyFaultActiveLastScan;
   Framework.AnyCriticalActive := Framework.AnyCriticalActiveLastScan;
   Framework.AnySimulationOn := Framework.AnySimulationOnLastScan;
   Framework.AnyHandOn := Framework.AnyHandOnLastScan;
   Framework.AlarmCount := Framework.TempAlarmCount;
   
   // Reset scratch
   Framework.AnyAudibleOnLastScan := 0;
   Framework.AnyAlarmActiveLastScan := 0;
   Framework.AnyWarningActiveLastScan := 0;
   Framework.AnyFaultActiveLastScan := 0;
   Framework.AnyCriticalActiveLastScan := 0;
   Framework.AnySimulationOnLastScan := 0;
   Framework.AnyHandOnLastScan := 0;
   Framework.TempAlarmCount := 0;
   
   // Constants
   Framework.AlwaysTrue := 1;
   Framework.AlwaysFalse := 0;
   
   // Random
   CMoRandom(fbRandom,Framework.LastRandomSeed);
   Framework.Random := fbRandom.Out;
   Framework.LastRandomSeed := fbRandom.NewSeed;
   
   // Ticks
   tmTick100ms.PRE := 100;
   tmTick100ms.TimerEnable := 1;
   TONR(tmTick100ms);
   Framework.Tick100ms := tmTick100ms.DN;
   IF tmTick100ms.DN THEN tmTick100ms.Reset := 1; TONR(tmTick100ms); tmTick100ms.Reset := 0; END_IF;
   
   tmTick1s.PRE := 1000;
   tmTick1s.TimerEnable := 1;
   TONR(tmTick1s);
   Framework.Tick1s := tmTick1s.DN;
   IF tmTick1s.DN THEN tmTick1s.Reset := 1; TONR(tmTick1s); tmTick1s.Reset := 0; END_IF;
   
   tmTick10s.PRE := 10000;
   tmTick10s.TimerEnable := 1;
   TONR(tmTick10s);
   Framework.Tick10s := tmTick10s.DN;
   IF tmTick10s.DN THEN tmTick10s.Reset := 1; TONR(tmTick10s); tmTick10s.Reset := 0; END_IF;
   
   // Blinkers
   tmBlink100ms.PRE := 100;
   tmBlink100ms.TimerEnable := 1;
   TONR(tmBlink100ms);
   IF tmBlink100ms.DN THEN bState100ms := NOT bState100ms; tmBlink100ms.Reset := 1; TONR(tmBlink100ms); tmBlink100ms.Reset := 0; END_IF;
   Framework.Blink100ms := bState100ms;
   
   tmBlink250ms.PRE := 250;
   tmBlink250ms.TimerEnable := 1;
   TONR(tmBlink250ms);
   IF tmBlink250ms.DN THEN bState250ms := NOT bState250ms; tmBlink250ms.Reset := 1; TONR(tmBlink250ms); tmBlink250ms.Reset := 0; END_IF;
   Framework.Blink250ms := bState250ms;
   
   tmBlink500ms.PRE := 500;
   tmBlink500ms.TimerEnable := 1;
   TONR(tmBlink500ms);
   IF tmBlink500ms.DN THEN bState500ms := NOT bState500ms; tmBlink500ms.Reset := 1; TONR(tmBlink500ms); tmBlink500ms.Reset := 0; END_IF;
   Framework.Blink500ms := bState500ms;
   
   tmBlink1s.PRE := 1000;
   tmBlink1s.TimerEnable := 1;
   TONR(tmBlink1s);
   IF tmBlink1s.DN THEN bState1s := NOT bState1s; tmBlink1s.Reset := 1; TONR(tmBlink1s); tmBlink1s.Reset := 0; END_IF;
   Framework.Blink1s := bState1s;
   
   tmBlink2s.PRE := 2000;
   tmBlink2s.TimerEnable := 1;
   TONR(tmBlink2s);
   IF tmBlink2s.DN THEN bState2s := NOT bState2s; tmBlink2s.Reset := 1; TONR(tmBlink2s); tmBlink2s.Reset := 0; END_IF;
   Framework.Blink2s := bState2s;
   
   // Free-running timer
   Framework.FreeRunningTimer := Framework.FreeRunningTimer + 1;
   
   // DateTime
   CMoGetLocalDateTime(fbGetLocal,Framework.CurrentLocalDateTime);
   CMoGetUTCDateTime(fbGetUTC,Framework.CurrentUTCDateTime);
   CMoDateTimeToString(fbLocalToStr,Framework.CurrentLocalDateTime,Framework.CurrentLocalString);
   CMoDateTimeToString(fbUTCToStr,Framework.CurrentUTCDateTime,Framework.CurrentUTCString);
END_ROUTINE
END_ADD_ON_INSTRUCTION

ADD_ON_INSTRUCTION CMoRandom   (* revision 1.0 *)
// Random Number Generator
// Help:
// Park-Miller LCG. Outputs REAL 0.0 to 1.0.
VAR_INPUT
   Seed : DINT := 48271; {required}   // Input seed value
END_VAR
VAR_OUTPUT
   Out : REAL; {access Read Only}   // Random number 0.0-1.0
   NewSeed : DINT; {access Read Only}   // Output seed for next call
END_VAR

ROUTINE Logic   (* structured text *)
   // =============================================================================
   // CMoRandom — Random Number Generator
   // CMo Library v1.0
   // =============================================================================
   // Park-Miller linear congruential generator.
   // Outputs a REAL between 0.0 and 1.0.
   //
   // Feed Seed from Framework.LastRandomSeed, write NewSeed back after call.
   // Called internally by CMoMainRuntime every scan.
   //
   // Usage:
   //   CMoRandom(fbRandom, Framework.LastRandomSeed);
   //   Framework.Random := fbRandom.Out;
   //   Framework.LastRandomSeed := fbRandom.NewSeed;
   // =============================================================================
   
   IF Seed <= 0 THEN
       Seed := 1;
   END_IF;
   NewSeed := (Seed MOD 127773) * 16807 - (Seed / 127773) * 2836;
   IF NewSeed <= 0 THEN
       NewSeed := NewSeed + 2147483647;
   END_IF;
   Out := NewSeed / 2147483647.0;
END_ROUTINE
END_ADD_ON_INSTRUCTION

PROGRAM MainProgram   (* main routine MainRoutine *)
VAR
   delta : CMoDateTime;
   deltaTime : DINT;
   DI_GuardClosed : CMoHALDigitalInput;
   DI_PartPresent : CMoHALDigitalInput;
   DO_MotorRun : CMoHALDigitalOutput;
   fbDiffTime : CMoDiffTime;
   fbGuardClosed : CMoDigitalInput;
   fbInterlock : CMoEvalInterlock;
   fbMainRuntime : CMoMainRuntime;
   fbMotorRun : CMoDigitalOutput;
   fbPartPresent : CMoDigitalInput;
   Framework : CMoFramework;
   Interlock_Motor : CMoInterlock;
   SimGuardClosed : BOOL;
   SimPartPresent : BOOL;
   storeTime1 : BOOL;
   storeTime2 : BOOL;
   Time1 : CMoDateTime;
   Time2 : CMoDateTime;
END_VAR

ROUTINE MainRoutine   (* structured text *)
   // Declare these as controller-scoped tags:
   //   Framework : CMoFramework
   //   DI_PartPresent : CMoHALDigitalInput
   //   DI_GuardClosed : CMoHALDigitalInput
   //   DO_MotorRun : CMoHALDigitalOutput
   //   Interlock_Motor : CMoInterlock
   //   fbMainRuntime : CMoMainRuntime
   //   fbPartPresent : CMoDigitalInput
   //   fbGuardClosed : CMoDigitalInput
   //   fbMotorRun : CMoDigitalOutput
   //   fbInterlock : CMoEvalInterlock
   //   SimPartPresent : BOOL
   //   SimGuardClosed : BOOL
   
   // Heartbeat: always first
   CMoMainRuntime(fbMainRuntime, Framework);
   
   // Enable simulation globally
   Framework.SimulationEnabled := 1;
   
   // --- Part Present sensor ---
   DI_PartPresent.EnableSimulation := 1;
   DI_PartPresent.SimInput := SimPartPresent;
   DI_PartPresent.Name := 'Part Present';
   
   CMoDigitalInput(fbPartPresent, DI_PartPresent,0 ,1,Framework);
   
   // --- Guard Door sensor ---
   DI_GuardClosed.EnableSimulation := 1;
   DI_GuardClosed.SimInput := SimGuardClosed;
   DI_GuardClosed.Name := 'Guard Closed';
   
   CMoDigitalInput(fbGuardClosed, DI_GuardClosed,0  ,1,Framework);
   
   // --- Interlock ---
   Interlock_Motor.PointCount := 2;
   Interlock_Motor.Condition[0] := DI_PartPresent.Value;
   Interlock_Motor.Condition[1] := DI_GuardClosed.Value;
   
   CMoEvalInterlock(fbInterlock, Interlock_Motor);
   
   // --- Business logic: .Value only ---
   DO_MotorRun.EnableSimulation := 1;
   DO_MotorRun.Value := Interlock_Motor.OK;
   DO_MotorRun.Name := 'Motor Run';
   
   CMoDigitalOutput(fbMotorRun, DO_MotorRun,1 ,Framework);
   
   if (storeTime1) then
   	COP(Framework.CurrentUTCDateTime,Time1,1);
   end_if;
   
   if (storeTime2) then
   	COP(Framework.CurrentUTCDateTime,Time2,1);
   end_if;
   
   CMoDiffTime(fbDiffTime,Time1,Time2,delta);
   
   deltaTime := fbDiffTime.TotalMicroseconds;
END_ROUTINE
END_PROGRAM
